FUNCTION "naut_DIV_LINT" : LINT
{ S7_Optimized_Access := 'TRUE' }
VERSION : 0.1
   VAR_INPUT
      A : LINT;
      B : LINT;
   END_VAR

BEGIN
	IF #B = 0 THEN
		#naut_DIV_LINT := 0;
	ELSE
		#naut_DIV_LINT := #A / #B;
	END_IF;
END_FUNCTION
